Fanuc KAREL source: KO00109.KL

PROGRAM KO00109
%NOLOCKGROUP
VAR
  A: REAL
  B: ARRAY[2] OF BYTE
  OUT: INTEGER
BEGIN
  A = 1
  B[1] = 2
  OUT = ATAN2(A, B[1])
END KO00109
